(* IEC 61131-3 sources: 2026_Projet_YGO_ExcavatriceDragage/CODE_BACKUP/CODE_20260904_AvantWeekendBackup_v0.6.34/H_TREUILS_BENNE/BENNE/_TYPES, 2 files *)

(* ---- ST_fbBucket_Config.st ---- *)
(* =======================================================================
   ⚙️ ST_fbBucket_Config — Configuration des offsets du benne
   ───────────────────────────────────────────────────────────────
   🎯 Rôle : Structure de paramétrage des décalages et anticipations benne
   📄 Doc métier : DOC/AF/AF_Partie-10_Fonction_Winch_v2.1.md
   ======================================================================= *)
TYPE ST_fbBucket_Config :
STRUCT
    OffsetOpenM        : REAL;                                        // Ecart M1/M2 en metres benne ouvert (m)
    OffsetCloseM       : REAL;                                        // Ecart M1/M2 en metres benne ferme (m)
    CoherenceLimitM    : REAL;                                        // Seuil de detection d'incoherence au boot (m)
    CloseAnticipationM : REAL := 1.0;                                 // Anticipation coupure commande fermeture (m) -- reglable IHM
    OpenAnticipationM  : REAL := 1.3;                                 // Anticipation coupure commande ouverture (m) -- reglable IHM
    JogSlowdownZoneM   : REAL := 1.0;                                 // Distance avant le point d'arret anticipe ou le jog unitaire M2 est force au palier 1 (m) -- reglable IHM
END_STRUCT
END_TYPE

(* ---- ST_fbBucket_State.st ---- *)
(* =======================================================================
   🚦 ST_fbBucket_State — État mémorisé et diagnostic du benne
   ───────────────────────────────────────────────────────────────
   🎯 Rôle : Structure d'état physique mémorisé et de diagnostic du benne
   📄 Doc métier : DOC/AF/AF_Partie-10_Fonction_Winch_v2.1.md
   ======================================================================= *)
TYPE ST_fbBucket_State :
STRUCT
    IsOpen          : BOOL;                                           // Benne ouvert memorise
    IsClosed        : BOOL;                                           // Benne ferme memorise
    TooOpen         : BOOL;                                           // Depassement ouverture (Delta < OffsetOpen - Tolerance)
    TooClosed       : BOOL;                                           // Depassement fermeture (Delta > OffsetClose + Tolerance)
    IsIntermediate  : BOOL;                                           // Position intermediaire (entre Ouvert et Ferme)
    LastPosM2Open   : REAL;                                           // Derniere position M2 memorisee ouvert (m)
    LastPosM2Close  : REAL;                                           // Derniere position M2 memorisee ferme (m)
    ActiveOffsetValid : BOOL;                                         // Validite offset actif calcule a jour (LIVE : exige puissance + BucketReferenced)
    BucketReferenced : BOOL;                                          // Reference benne PERSISTANTE (RETAIN) : offsets calibres + datum M1/M2 fiables lors de la calibration. Survit a une coupure puissance. Retombe si M1/M2 suspect/incoherent, CfgFault, ou recalibration explicite.
    StateIncoherent : BOOL;                                           // Etat non sur (divergence boot/reel)
END_STRUCT
END_TYPE
